Staubli VAL3: default.pjx

--- default.pjx ---
parameters version=s6.8 stackSize=5000 millimeterUnit=true
program file=start.pgx
program file=stop.pgx
data file=default.dtx
alias name=io interface=io autoload=true password=

--- default.dtx ---


--- start.pgx ---
program start()
begin
end

--- stop.pgx ---
program stop()
begin
end
